# EPICS substitutions: 1.5.0/debian-12/7.0.10/base/templates/makeBaseApp/top/exampleApp/Db/user.substitutions
# SPDX-FileCopyrightText: 2006 Argonne National Laboratory
#
# SPDX-License-Identifier: EPICS

# Example substitutions file

file "db/circle.db" {
    { user = "_USER_" }
}

file "db/dbExample1.db" {
    { user = "_USER_" }
}

file db/dbExample2.db {
    pattern { user, no, scan }
        { "_USER_", 1, "1 second" }
        { "_USER_", 2, "2 second" }
        { "_USER_", 3, "5 second" }
}
